Fanuc KAREL source: KA00165.KL

PROGRAM KA00165
%NOLOCKGROUP
VAR
  SRC: ARRAY[4] OF BOOLEAN
  DST: ARRAY[4] OF BOOLEAN
BEGIN
  DST = SRC
END KA00165
